(* PLC project Pumps.project, CODESYS CODESYS V3.5 SP19 *)
(* stored: creationDateTime 2026-10-22T10:00:00, modificationDateTime 2026-10-22T10:00:00 *)

FUNCTION Il_Limit : INT
  VAR_INPUT
    nIn : INT;
    nMax : INT;
  END_VAR

            LD   nIn
GT   nMax     (* above the limit? *)
JMPC Clip
LD   nIn
ST   Il_Limit
RET
Clip:
LD   nMax
ST   Il_Limit
          
END_FUNCTION

PROGRAM Cfc_Pump
  VAR
    bRun : BOOL;
    bOk : BOOL;
    bMotor : BOOL;
  END_VAR

(* CFC diagram, written out as Structured Text *)
END_PROGRAM
